(* IEC 61131-3 sources: Industry-PLC-LLM/data/PLCBEAD_repo/PLCBEAD_PLCEmbed-main/PLC-BEAD/Source/PLC_Programs (part 16) *)

(* ---- UTC_TO_LTIME.ST ---- *)
FUNCTION _INT_TO_UDINT:UDINT
	VAR_INPUT
		IN :	INT;
	END_VAR

	_INT_TO_UDINT := DINT_TO_UDINT(INT_TO_DINT(IN));
END_FUNCTION

FUNCTION DT_TO_DATE2:UDINT
	VAR_INPUT
		IN :	UDINT;
	END_VAR

	DT_TO_DATE2 := (IN / UDINT#86400) * UDINT#86400;
END_FUNCTION

FUNCTION YEAR_OF_DATE:INT
	VAR_INPUT
		IDATE :	UDINT;
	END_VAR

	YEAR_OF_DATE := UDINT_TO_INT((idate+UDINT#43200) / UDINT#31557600 + UDINT#1970);
END_FUNCTION

FUNCTION SET_DT:UDINT

	VAR_INPUT
		YEAR : INT;
		MONTH :	INT;
		DAY : INT;
		HOUR : INT;
		MINUTE : INT;
		SECOND : INT;
	END_VAR

	SET_DT := SET_DATE(YEAR, MONTH, DAY) + _INT_TO_UDINT(SECOND) + _INT_TO_UDINT(MINUTE) * UDINT#60 + _INT_TO_UDINT(HOUR) * UDINT#3600;

END_FUNCTION

FUNCTION SET_DATE:UDINT

	VAR_INPUT
		YEAR :	INT;
		MONTH :	INT;
		DAY :	INT;
	END_VAR

	VAR
		count :	INT;
	END_VAR

	IF month > 2 THEN
		count := (month - 1) * 30;
		IF month > 7 THEN
			count := count + DWORD_TO_INT(SHR(DINT_TO_DWORD(INT_TO_DINT(month) - INT_TO_DINT(3)),1));
		ELSE
			count := count + DWORD_TO_INT(SHR(DINT_TO_DWORD(INT_TO_DINT(month) - INT_TO_DINT(4)),1));
		END_IF;
		IF SHL(INT_TO_WORD(year),14) = WORD#0 THEN
			count := count + 1;
		END_IF;
	ELSE
		count := (month - 1) * 31;
	END_IF;
	SET_DATE := (_INT_TO_UDINT(count + day - 1) + DWORD_TO_UDINT(SHR(UDINT_TO_DWORD(_INT_TO_UDINT(year) * UDINT#1461 - UDINT#2878169), 2))) * UDINT#86400;

END_FUNCTION

FUNCTION DST:BOOL
	VAR_INPUT
		UTC :	UDINT;
	END_VAR

	VAR
		yr :	INT;
		yr4 :	UDINT;
		ltc :	UDINT;
		idate :	UDINT;
	END_VAR

	yr := YEAR_OF_DATE(DT_TO_DATE2(UTC));
	ltc := UTC;
	idate := SET_DT(yr, 3, 31, 1, 0, 0);
	yr4 := DWORD_TO_UDINT(SHR(INT_TO_DWORD(5 * yr), 2)) + UDINT#1;
	DST := (idate - ((yr4 + UDINT#3) MOD UDINT#7) * UDINT#86400 <= ltc) AND (idate + (UDINT#214 - (yr4) MOD UDINT#7) * UDINT#86400 > ltc);

END_FUNCTION

FUNCTION UTC_TO_LTIME:UDINT

	VAR_INPUT
		UTC :	UDINT;
		DST_ENABLE :	BOOL;
		TIME_ZONE_OFFSET :	INT;
	END_VAR

	VAR
		tmp :	INT;
	END_VAR

	UTC_TO_LTIME := UTC + _INT_TO_UDINT(TIME_ZONE_OFFSET) * UDINT#60 + BOOL_TO_UDINT(DST_ENABLE AND DST(UTC)) * UDINT#3600;

	tmp := TIME_ZONE_OFFSET * 60 + BOOL_TO_INT(DST_ENABLE AND DST(UTC)) * 3600;
	IF tmp < 0 THEN
		UTC_TO_LTIME := UTC - _INT_TO_UDINT(ABS(tmp));
	ELSE
		UTC_TO_LTIME := UTC + _INT_TO_UDINT(tmp);
	END_IF;

END_FUNCTION

PROGRAM program0
  VAR
	UTC :	UDINT;
	DST_ENABLE :	BOOL;
	TIME_ZONE_OFFSET :	INT;
    CEIL5_OUT : UDINT;
  END_VAR

  CEIL5_OUT := UTC_TO_LTIME(UTC, DST_ENABLE, TIME_ZONE_OFFSET);
END_PROGRAM

CONFIGURATION Config0

  RESOURCE Res0 ON PLC
    TASK task0(INTERVAL := T#20ms,PRIORITY := 0);
    PROGRAM instance0 WITH task0 : program0;
  END_RESOURCE
END_CONFIGURATION

(* ---- WATER_DENSITY.ST ---- *)
FUNCTION WATER_DENSITY:REAL

    VAR_INPUT
        T :	REAL;
        SAT :	BOOL;
    END_VAR

    VAR
        T2 :	REAL;
        T4 :	REAL;
    END_VAR

    T2 := T * T;
    T4 := T2 * T2;
    WATER_DENSITY := (999.83952 + 16.952577*T + -7.9905127E-3*T2 + -4.6241757E-5*T2*T + 1.0584601E-7*T4 + -2.8103006E-10*T4*T) / (1.0 + 0.0168872*T);
    IF sat THEN WATER_DENSITY := WATER_DENSITY - 0.004612 + 0.000106 * T; END_IF;

END_FUNCTION

PROGRAM program0
	VAR
		T :	REAL;
        SAT :	BOOL;
		CEIL5_OUT : REAL;
	END_VAR

  	CEIL5_OUT := WATER_DENSITY(T, SAT);
END_PROGRAM

CONFIGURATION Config0

  RESOURCE Res0 ON PLC
    TASK task0(INTERVAL := T#20ms,PRIORITY := 0);
    PROGRAM instance0 WITH task0 : program0;
  END_RESOURCE
END_CONFIGURATION

(* ---- WCT.ST ---- *)
FUNCTION WCT:REAL

	VAR_INPUT
		T :	REAL;
		V :	REAL;
	END_VAR

	IF V < 5.0 OR T > 10.0 THEN
		WCT := T;
	ELSE
		WCT := 13.12 + 0.6215 * T +(0.3965 * T - 11.37) * EXP(LN(v) * 0.16);
	END_IF;

END_FUNCTION

PROGRAM program0
	VAR
		T :	REAL;
		V :	REAL;
		CEIL5_OUT : REAL;
	END_VAR

  	CEIL5_OUT := WCT(T, V);
END_PROGRAM

CONFIGURATION Config0

  RESOURCE Res0 ON PLC
    TASK task0(INTERVAL := T#20ms,PRIORITY := 0);
    PROGRAM instance0 WITH task0 : program0;
  END_RESOURCE
END_CONFIGURATION

(* ---- WINDOW.ST ---- *)
FUNCTION WINDOW:BOOL
	VAR_INPUT
		LOW :	REAL;
		IN :	REAL;
		HIGH :	REAL;
	END_VAR
	window := (in < high) AND (in > low);

END_FUNCTION

PROGRAM program0
  	VAR
		LOW :	REAL;
		IN :	REAL;
		HIGH :	REAL;
		CEIL5_OUT : BOOL;
	END_VAR

  	CEIL5_OUT := window(LOW, IN, HIGH);
END_PROGRAM

CONFIGURATION Config0
  	RESOURCE Res0 ON PLC
    	TASK task0(INTERVAL := T#20ms,PRIORITY := 0);
    	PROGRAM instance0 WITH task0 : program0;
  	END_RESOURCE
END_CONFIGURATION

(* ---- WINDOW2.ST ---- *)
FUNCTION WINDOW2:BOOL
	VAR_INPUT
		LOW :	REAL;
		IN :	REAL;
		HIGH :	REAL;
	END_VAR
	window2 := (in <= high) AND (in >= low);
END_FUNCTION

PROGRAM program0
  	VAR
		LOW :	REAL;
		IN :	REAL;
		HIGH :	REAL;
		CEIL5_OUT : BOOL;
	END_VAR

  	CEIL5_OUT := window2(LOW, IN, HIGH);
END_PROGRAM

CONFIGURATION Config0
  	RESOURCE Res0 ON PLC
    	TASK task0(INTERVAL := T#20ms,PRIORITY := 0);
    	PROGRAM instance0 WITH task0 : program0;
  	END_RESOURCE
END_CONFIGURATION

(* ---- WORD_OF_BYTE.ST ---- *)
FUNCTION WORD_OF_BYTE:WORD
	VAR_INPUT
		B1 :	BYTE;
		B0 :	BYTE;
	END_VAR
	WORD_OF_BYTE := SHL(BYTE_TO_WORD(B1),8) OR BYTE_TO_WORD(B0);
END_FUNCTION

PROGRAM program0
  	VAR
		B1 :	BYTE;
		B0 :	BYTE;
		CEIL5_OUT : WORD;
	END_VAR

  	CEIL5_OUT := WORD_OF_BYTE(B1, B0);
END_PROGRAM

CONFIGURATION Config0
  	RESOURCE Res0 ON PLC
    	TASK task0(INTERVAL := T#20ms,PRIORITY := 0);
    	PROGRAM instance0 WITH task0 : program0;
  	END_RESOURCE
END_CONFIGURATION

(* ---- WORD_OF_DWORD.ST ---- *)
FUNCTION _BYTE_TO_INT:INT
	VAR_INPUT
		IN :	BYTE;
	END_VAR

	_BYTE_TO_INT := USINT_TO_INT(BYTE_TO_USINT(IN));
END_FUNCTION

FUNCTION WORD_OF_DWORD:WORD
	VAR_INPUT
		IN: DWORD;
		N :	BYTE;
	END_VAR
	WORD_OF_DWORD := DWORD_TO_WORD(SHR(in,_BYTE_TO_INT(SHL(n,4))));
END_FUNCTION

PROGRAM program0
  	VAR
		IN :	DWORD;
		N :	BYTE;
		CEIL5_OUT : WORD;
	  END_VAR

  	CEIL5_OUT := WORD_OF_DWORD(IN, N);
END_PROGRAM

CONFIGURATION Config0
  	RESOURCE Res0 ON PLC
    	TASK task0(INTERVAL := T#20ms,PRIORITY := 0);
    	PROGRAM instance0 WITH task0 : program0;
  	END_RESOURCE
END_CONFIGURATION

(* ---- WORD_TO_RANGE.ST ---- *)
FUNCTION _WORD_TO_REAL:REAL
	VAR_INPUT
		IN :	WORD;
	END_VAR
	_WORD_TO_REAL := UINT_TO_REAL(WORD_TO_UINT(IN));
END_FUNCTION

FUNCTION WORD_TO_RANGE:REAL
	VAR_INPUT
		X :	WORD;
		LOW :	REAL;
		HIGH :	REAL;
	END_VAR
	WORD_TO_RANGE := (high - low) * _WORD_TO_REAL(X) * 0.00001525902189669640 + low;
END_FUNCTION

PROGRAM program0
  	VAR
		X :	WORD;
		LOW :	REAL;
		HIGH :	REAL;
		CEIL5_OUT : REAL;
	  END_VAR

  	CEIL5_OUT := WORD_TO_RANGE(X, LOW, HIGH);
END_PROGRAM

CONFIGURATION Config0
  	RESOURCE Res0 ON PLC
    	TASK task0(INTERVAL := T#20ms,PRIORITY := 0);
    	PROGRAM instance0 WITH task0 : program0;
  	END_RESOURCE
END_CONFIGURATION

(* ---- WORK_WEEK.ST ---- *)
FUNCTION LEAP_YEAR:BOOL

  VAR_INPUT
    YEAR :	INT;
  END_VAR

  IF (year MOD INT#400) = INT#00 THEN
    leap_year := TRUE;
  ELSIF (year MOD INT#100) = INT#00 THEN
    leap_year := FALSE;
  ELSIF (year MOD INT#04) = INT#00 THEN
    leap_year := TRUE;
  ELSE
    leap_year := FALSE;
  END_IF;

END_FUNCTION

FUNCTION DAY_OF_WEEK:INT

	VAR_INPUT
		IDATE :	UDINT;
	END_VAR

	DAY_OF_WEEK := UDINT_TO_INT((idate / UDINT#86400 + UDINT#3) MOD UDINT#7) + INT#01;

END_FUNCTION

FUNCTION YEAR_OF_DATE:INT
	VAR_INPUT
		IDATE :	UDINT;
	END_VAR

	YEAR_OF_DATE := UDINT_TO_INT((idate+UDINT#43200) / UDINT#31557600 + UDINT#1970);
END_FUNCTION

FUNCTION _INT_TO_UDINT:UDINT
	VAR_INPUT
		IN :	INT;
	END_VAR

	_INT_TO_UDINT := DINT_TO_UDINT(INT_TO_DINT(IN));
END_FUNCTION

FUNCTION YEAR_BEGIN:UDINT
	VAR_INPUT
		Y :	INT;
	END_VAR
	year_begin := DWORD_TO_UDINT(SHR(UDINT_TO_DWORD(_INT_TO_UDINT(y) * UDINT#1461 - UDINT#2878169),2))*UDINT#86400;

END_FUNCTION

FUNCTION WORK_WEEK:INT

	VAR_INPUT
		IDATE :	UDINT;
	END_VAR

	VAR
		d1 :	UDINT;
		w1 :	INT;
		ds :	UDINT;
		yr :	INT;
		w31 :	INT;
		w01 :	INT;
		wm :	INT;
	END_VAR

	yr := YEAR_OF_DATE(idate);
	d1 := year_begin(yr);
	w1 := DAY_OF_WEEK(d1);
	IF w1 < 5 THEN
		ds := d1 - _INT_TO_UDINT(w1+6) * UDINT#86400;
	ELSE
		ds := d1 + _INT_TO_UDINT(1-w1) * UDINT#86400;
	END_IF;

	work_week := UDINT_TO_INT((idate - ds) / UDINT#604800);

	IF work_week = 0 THEN
		IF w1 > 1 THEN w31 := w1 - 1; ELSE W31 := 7; END_IF;
		IF leap_year(yr - 1) THEN IF w31 > 1 THEN w01 := W31 - 1; ELSE w1 := 7; END_IF; END_IF;
		WORK_WEEK := 52 + BOOL_TO_INT(w31 = 4 OR w01 = 4);
	ELSE
		IF leap_year(yr) THEN
			IF w1 < 7 THEN w31 := w1 + 1; ELSE w31 := 1; END_IF;
		ELSE
			w31 := w1;
		END_IF;
		wm := 52 + BOOL_TO_INT(w31 = 4 OR w1 = 4);
		IF work_week > wm THEN work_week := 1; END_IF;
	END_IF;

END_FUNCTION

PROGRAM program0
  VAR
    Y : UDINT;
    CEIL5_OUT : INT;
  END_VAR

  CEIL5_OUT := WORK_WEEK(Y);
END_PROGRAM

CONFIGURATION Config0

  RESOURCE Res0 ON PLC
    TASK task0(INTERVAL := T#20ms,PRIORITY := 0);
    PROGRAM instance0 WITH task0 : program0;
  END_RESOURCE
END_CONFIGURATION
